// TIA Portal V20 export
// export: Created 2026-10-20T18:55:00.357363Z, ExportSetting None, DisplayName Totally Integrated Automation Portal, DisplayVersion V20 Update 6, DisplayName TIA Portal Openness, DisplayVersion V20 Update 6, DisplayName TIA Portal Version Control Interface, DisplayVersion V20 Update 6, DisplayName SINAMICS Startdrive Advanced, DisplayVersion V20 SP1, DisplayName SINAMICS Startdrive G130, G150, S120, S150, SINAMICS MV, G220, S200, S210, DisplayVersion V20 SP1, DisplayName SINAMICS Startdrive G110M, G120, G120C, G120D, G120P, G115D, DisplayVersion V20 SP1, DisplayName STEP 7 Professional, DisplayVersion V20 Update 6, DisplayName STEP 7 Safety, DisplayVersion V20 Update 2, DisplayName WinCC Basic/Comfort/Advanced, DisplayVersion V20 Update 6, DisplayName WinCC Unified, DisplayVersion V20 Update 6
VAR_GLOBAL   // PLC tag table "IO_Remote_Panel_3"
   "Power Enable Safety Stopper Conveyors (Level 7,8 - Side1) - CH1(3)" AT %Q786.0 : Bool;
   "Power Enable Safety Stopper Conveyors (Level 7,8 - Side1) - CH2(3)" AT %Q786.1 : Bool;
   "Power Enable Safety Stopper Conveyors (Level 7,8 - Side2) - CH1(3)" AT %Q786.2 : Bool;
   "Power Enable Safety Stopper Conveyors (Level 7,8 - Side2) - CH2(3)" AT %Q786.3 : Bool;
   "VTU HOIST BRAKE SAFETY ENABLE 1(3)" AT %Q786.4 : Bool;
   "VTU HOIST BRAKE SAFETY ENABLE 2(3)" AT %Q786.5 : Bool;
   "Power Enable Safety Stopper Conveyors (Level 1,2,3 - Side2) - CH1(3)" AT %Q780.2 : Bool;
   "Power Enable Safety Stopper Conveyors (Level 1,2,3 - Side2) - CH2(3)" AT %Q780.3 : Bool;
   "Power Enable Safety Stopper Conveyors (Level 4,5,6 - Side2) - CH1(3)" AT %Q780.6 : Bool;
   "Power Enable Safety Stopper Conveyors (Level 4,5,6 - Side2) - CH2(3)" AT %Q780.7 : Bool;
   "STO CNV VFD (Level 1,2,3 - Side2) - CH1(3)" AT %Q768.6 : Bool;
   "STO CNV VFD (Level 1,2,3 - Side2) - CH2(3)" AT %Q768.7 : Bool;
   "STO CNV VFD (Level 4,5,6 - Side1) - CH1(3)" AT %Q774.0 : Bool;
   "STO CNV VFD (Level 4,5,6 - Side1) - CH2(3)" AT %Q774.1 : Bool;
   "STO CNV VFD (Level 4,5,6 - Side2) - CH1(3)" AT %Q774.2 : Bool;
   "STO CNV VFD (Level 4,5,6 - Side2) - CH2(3)" AT %Q774.3 : Bool;
   "STO CNV VFD (Level 7,8 - Side1) - CH1(3)" AT %Q774.4 : Bool;
   "STO CNV VFD (Level 7,8 - Side1) - CH2(3)" AT %Q774.5 : Bool;
   "STO CNV VFD (Level 7,8 - Side2) - CH1(3)" AT %Q774.6 : Bool;
   "STO CNV VFD (Level 7,8 - Side2) - CH2(3)" AT %Q774.7 : Bool;
   "VTD3 PUSH TO EXIT VTD ZONE" AT %I363.5 : Bool;
   "Power Enable Safety Stopper Conveyors (Level 1,2,3 - Side1) - CH2(3)" AT %Q780.1 : Bool;
   "STO CONVEYOR VTD - CH1(3)" AT %Q768.2 : Bool;
   "RESET (CABINET)(3)" AT %I740.3 : Bool;   // Reset (Cabinet) - CH1
   "STO VTD - CH2(3)" AT %Q768.1 : Bool;
   "STO VTD - CH1(3)" AT %Q768.0 : Bool;
   "STO CNV VFD (Level 1,2,3 - Side1) - CH1(3)" AT %Q768.4 : Bool;
   "STO CONVEYOR VTD - CH2(3)" AT %Q768.3 : Bool;
   "CABINET 24V PSU CIRCUIT BREAKER FEEDBACK(3)" AT %I366.2 : Bool;
   "VTD3 CIRCUIT BREAKER FEEDBACK" AT %I366.1 : Bool;
   "VTD3 PUSH TO ENTER VTD ZONE" AT %I363.4 : Bool;
   "OVERTRAVEL UPPER LIMIT - CH2(3)" AT %I740.5 : Bool;   // Overtravel Upper Limit - CH2
   "Power Enable Safety Stopper Conveyors (Level 1,2,3 - Side1) - CH1(3)" AT %Q780.0 : Bool;
   "CABINET COOLING FAN CIRCUIT BREAKER FEEDBACK(3)" AT %I366.3 : Bool;
   "STO CNV VFD (Level 1,2,3 - Side1) - CH2(3)" AT %Q768.5 : Bool;
   "VTD3 LOWER LIMIT" AT %I362.3 : Bool;
   "VTD3 UPPER LIMIT" AT %I362.0 : Bool;
   "OVERTRAVEL LOWER LIMIT - CH2(3)" AT %I740.4 : Bool;   // Overtravel Lower Limit - CH2
   "Power Enable Safety Stopper Conveyors (Level 4,5,6 - Side1) - CH1(3)" AT %Q780.4 : Bool;
   "E-STOP (CABINET) - CH2(3)" AT %I740.6 : Bool;   // E-Stop (Cabinet) - CH2
   "OVERTRAVEL LOWER LIMIT - CH1(3)" AT %I740.0 : Bool;   // Overtravel Lower Limit - CH1
   "Power Enable Safety Stopper Conveyors (Level 4,5,6 - Side1) - CH2(3)" AT %Q780.5 : Bool;
   "OVERTRAVEL UPPER LIMIT - CH1(3)" AT %I740.1 : Bool;   // Overtravel Upper Limit - CH1
   "E-STOP (CABINET) - CH1(3)" AT %I740.2 : Bool;   // E-Stop (Cabinet)- CH1
   "CVTD3 CIRCUIT BREAKER FEEDBACK" AT %I366.0 : Bool;
   "EMERGENCY STOP RESET STATUS - ON(3)" AT %Q484.7 : Bool;   // 920SL1
   "VTD3 SFTY STOPPER CNVS 7,8 - (SIDE 2)" AT %I754.5 : Bool;
   "VTU HOIST BRAKE SAFETY ENABLE EDM FEEDBACK(3)" AT %I754.6 : Bool;
   "VTD3 SFTY STOPPER CNVS 4,5,6 - (SIDE 1)" AT %I754.2 : Bool;
   "VTD3 SFTY STOPPER CNVS 7,8 - (SIDE 1)" AT %I754.4 : Bool;
   "VTD3 SFTY STOPPER CNVS 4,5,6 - (SIDE 2)" AT %I754.3 : Bool;
   "VTD3 SFTY STOPPER CNVS 1,2,3 - (SIDE 2)" AT %I754.1 : Bool;
   "VTD3 SFTY STOPPER CNVS 1,2,3 - (SIDE 1)" AT %I754.0 : Bool;   // SAFETY STOPPER CONVEYORS (1,2,3 - SIDE 1) EDMFEEDBACK
   "C3107 CIRCUIT BREAKER FEEDBACK" AT %I365.6 : Bool;
   "C3204 CIRCUIT BREAKER FEEDBACK" AT %I364.3 : Bool;
   "C3102 CIRCUIT BREAKER FEEDBACK" AT %I365.1 : Bool;
   "C3105 CIRCUIT BREAKER FEEDBACK" AT %I365.4 : Bool;
   "C3203 CIRCUIT BREAKER FEEDBACK" AT %I364.2 : Bool;
   "C3106 CIRCUIT BREAKER FEEDBACK" AT %I365.5 : Bool;
   "C3208 CIRCUIT BREAKER FEEDBACK" AT %I364.7 : Bool;
   "C3205 CIRCUIT BREAKER FEEDBACK" AT %I364.4 : Bool;
   "C3101 CIRCUIT BREAKER FEEDBACK" AT %I365.0 : Bool;
   "C3108 CIRCUIT BREAKER FEEDBACK" AT %I365.7 : Bool;
   "Chain Slack 3 - CH1(3)" AT %I747.1 : Bool;   // Chain Slack 3 - CH1
   "Chain Slack 4 - CH1(3)" AT %I747.0 : Bool;   // Chain Slack 4 - CH1
   "Chain Slack 1 - CH2(3)" AT %I747.7 : Bool;   // Chain Slack 1 - CH2
   "C3103 CIRCUIT BREAKER FEEDBACK" AT %I365.2 : Bool;
   "Chain Slack 1 - CH1(3)" AT %I747.3 : Bool;   // Chain Slack 1 - CH1
   "Chain Slack 2 - CH1(3)" AT %I747.2 : Bool;   // Chain Slack 2 - CH1
   "C3104 CIRCUIT BREAKER FEEDBACK" AT %I365.3 : Bool;
   "SCA 3002 STACK LIGHTS ORANGE" AT %Q484.5 : Bool;
   "C3202 CIRCUIT BREAKER FEEDBACK" AT %I364.1 : Bool;
   "Chain Slack 3 - CH2(3)" AT %I747.5 : Bool;   // Chain Slack 3 - CH2
   "SCA 3002 STACK LIGHTS RED" AT %Q484.4 : Bool;
   "Chain Slack 2 - CH2(3)" AT %I747.6 : Bool;   // Chain Slack 2 - CH2
   "Chain Slack 4 - CH2(3)" AT %I747.4 : Bool;   // Chain Slack 4 - CH2
   "C3206 CIRCUIT BREAKER FEEDBACK" AT %I364.5 : Bool;
   "C3201 CIRCUIT BREAKER FEEDBACK" AT %I364.0 : Bool;
   "SCA 3002 STACK LIGHTS GREEN" AT %Q484.6 : Bool;
   "C3207 CIRCUIT BREAKER FEEDBACK" AT %I364.6 : Bool;
   "C3105_SFTY STOPPER ROTATE" AT %Q482.0 : Bool;
   "C3107_SFTY STOPPER ROTATE" AT %Q483.0 : Bool;
   "C3206_SFTY STOPPER ROTATE" AT %Q478.4 : Bool;
   "C3103_SFTY STOPPER ROTATE" AT %Q481.0 : Bool;
   "C3203_SFTY STOPPER ROTATE" AT %Q477.0 : Bool;
   "C3108_SFTY STOPPER ROTATE" AT %Q483.4 : Bool;
   "C3106_SFTY STOPPER ROTATE" AT %Q482.4 : Bool;
   "C3207_SFTY STOPPER ROTATE" AT %Q479.0 : Bool;
   "C3202_SFTY STOPPER ROTATE" AT %Q476.4 : Bool;
   "C3204_SFTY STOPPER ROTATE" AT %Q477.4 : Bool;
   "C3101_SFTY STOPPER ROTATE" AT %Q480.0 : Bool;
   "C3208_SFTY STOPPER ROTATE" AT %Q479.4 : Bool;
   "C3201_SFTY STOPPER ROTATE" AT %Q476.0 : Bool;
   "C3205_SFTY STOPPER ROTATE" AT %Q478.0 : Bool;
   "C3102_SFTY STOPPER ROTATE" AT %Q481.4 : Bool;
   "C3104_SFTY STOPPER ROTATE" AT %Q480.4 : Bool;
   "LIGHT GUARDS C3101 - CH2" AT %I761.5 : Bool;
   "LIGHT GUARDS C3201 - CH1" AT %I761.0 : Bool;
   "LIGHT GUARDS C3201 - CH2" AT %I761.4 : Bool;
   "LIGHT GUARDS C3101 - CH1" AT %I761.1 : Bool;
   "VTD3 DOCKING PINS 1 EXTEND" AT %Q484.0 : Bool;
   "VTD3 DOCKING PINS 2 RETRACT" AT %Q484.3 : Bool;
   "VTD3 DOCKING PINS 1 RETRACT" AT %Q484.1 : Bool;
   "VTD3 DOCKING PINS 2 EXTEND" AT %Q484.2 : Bool;
   "GATE_SENSOR_1_CH2(3)" AT %I761.7 : Bool;
   "GATE_SENSOR_2_CH1(3)" AT %I761.2 : Bool;
   "GATE_SENSOR_2_CH2(3)" AT %I761.6 : Bool;
   "GATE_SENSOR_1_CH1(3)" AT %I761.3 : Bool;
END_VAR
